SUBAPPLICATION logiBUS_AI_Calibrate_2P_IDA_Param_OPC (* logiBUS_AI_IDA (Analog-Eingang) mit 2-Punkt-Kalibrierung (AR_CALIBRATE_2P_REF, unabhaengig gespeicherte Rohwerte X_LOW/X_HIGH + Referenzwerte LOW_REF/HIGH_REF alle INI-persistiert) auf VT-Zahlenfelder (Rohwert + kalibrierter Wert, je eigene CNumberVariable) + Bargraph (kalibriert) + 2 VT-Tasten (CO/CS) + OPC-UA (Rohwert DWORD + kalibrierter Wert REAL, generisch, ein Kanal) *)
  (* Standard: 61499-2; Description: Copyright (c) 2026 Meisterschulen am Ostbahnhof This program and the accompanying materials are made available under the terms of the Eclipse Public License 2.0 which is available at https://www.eclipse.org/legal/epl-2.0/ SPDX-License-Identifier: EPL-2.0 *)
  (* Version 1.0, 2026-11-23, Franz Höpfinger, Meisterschulen am Ostbahnhof, Kopie von logiBUS_AI_Calibrate_2P_IDA_OPC (v1.13), InputRaw jetzt logiBUS_AI_Raw_VT_AR_Param_OPC: Hysterese/TimeDelta/TimeRateLimit des AI per Web + INI einstellbar (gleiche sSection). Zuerst fuer Ultraschall B01. PublishCal auf AR_TO_Q_Publish_Fast_OPC: CAL-Publish ungedrosselt, nur VT-Anzeige 500 ms. *)
  PACKAGE MyLib::sys;
  IMPORT isobus::UT::Q::const::IDs::ID_NULL;
  IMPORT logiBUS::io::AI::logiBUS_AI;
  IMPORT logiBUS::io::AI::logiBUS_AI_S;
  IMPORT logiBUS::utils::conversion::phys::NumericObjectPool_S;
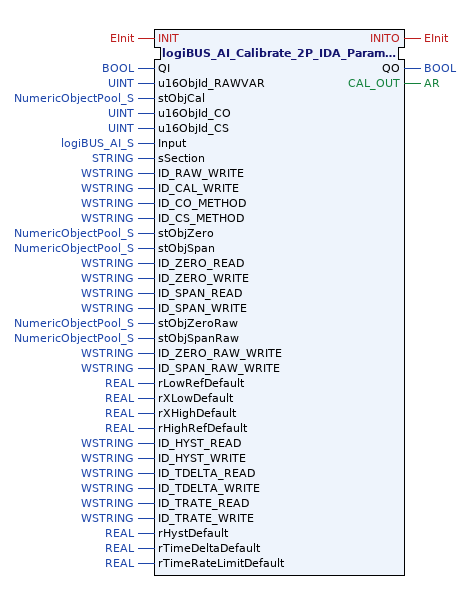
  EVENT_INPUT
    INIT : EInit; (* Initialization Request *)
  END_EVENT
  EVENT_OUTPUT
    INITO : EInit; (* Initialization Confirm *)
  END_EVENT
  VAR_INPUT
    QI : BOOL := TRUE; (* Quality Input - TRUE to enable service *)
    u16ObjId_RAWVAR : UINT := ID_NULL; (* Object ID CNumberVariable (Rohwert 0-4095, unkalibriert, reine Diagnose-Anzeige) *)
    stObjCal : logiBUS::utils::conversion::phys::NumericObjectPool_S := (u16ObjId := ID_NULL, r32Scale := 1.0, i32Offset := 0, u8Decimals := 1); (* Object ID + Scale/Offset/Decimals CNumberVariable (kalibrierter Wert, eigene, unabhaengige CNumberVariable) *)
    u16ObjId_CO : UINT := ID_NULL; (* Object ID Taste 'CO' (Kalibrier-Nullpunkt: Referenz 1 anlegen, dann druecken) *)
    u16ObjId_CS : UINT := ID_NULL; (* Object ID Taste 'CS' (Kalibrier-Spanne: Referenz 2 anlegen, dann druecken - erst nach CO moeglich) *)
    Input : logiBUS::io::AI::logiBUS_AI_S := logiBUS_AI::Invalid; (* Identify the Input AnalogInput_I1..I8 *)
    sSection : STRING; (* INI-Sektionsname fuer OFFSET/SCALE-Persistenz - pro Kanal eindeutig (z.B. 'AI_Calibrate_I1'), sonst kollidieren die Kanaele in settings.ini *)
    ID_RAW_WRITE : WSTRING; (* Rohwert-Ruckmelde-Adresse (DWORD 0-4095, ACTION=PUBLISH) *)
    ID_CAL_WRITE : WSTRING; (* Kalibrierter-Wert-Ruckmelde-Adresse (REAL, ACTION=PUBLISH) *)
    ID_CO_METHOD : WSTRING; (* Methodenadresse (ACTION=CREATE_METHOD) fuer den argumentlosen CO-Trigger - gleichberechtigt zur lokalen VT-Taste aufrufbar, sowohl vom OPC-UA-Dashboard als auch per CLIENT_0 von einer anderen Station (Cross-Station-Weiterleitung einer dortigen VT-Taste, siehe OPC_UA_VERNETZUNG.md Punkt 14 - kein Toggle/Subscribe-Umweg mehr) *)
    ID_CS_METHOD : WSTRING; (* Methodenadresse (ACTION=CREATE_METHOD) fuer den argumentlosen CS-Trigger - siehe ID_CO_METHOD *)
    stObjZero : logiBUS::utils::conversion::phys::NumericObjectPool_S := (u16ObjId := ID_NULL, r32Scale := 1.0, i32Offset := 0, u8Decimals := 1); (* Object ID + Scale/Offset/Decimals CNumberVariable (ZERO-Referenzwert, VT-Eingabefeld + OPC-UA) *)
    stObjSpan : logiBUS::utils::conversion::phys::NumericObjectPool_S := (u16ObjId := ID_NULL, r32Scale := 1.0, i32Offset := 0, u8Decimals := 1); (* Object ID + Scale/Offset/Decimals CNumberVariable (SPAN-Referenzwert, VT-Eingabefeld + OPC-UA) *)
    ID_ZERO_READ : WSTRING; (* Remote-Subscribe-Adresse ZERO-Referenzwert (REAL, ACTION=SUBSCRIBE) *)
    ID_ZERO_WRITE : WSTRING; (* Remote-Echo-Adresse ZERO-Referenzwert (REAL, ACTION=PUBLISH) *)
    ID_SPAN_READ : WSTRING; (* Remote-Subscribe-Adresse SPAN-Referenzwert (REAL, ACTION=SUBSCRIBE) *)
    ID_SPAN_WRITE : WSTRING; (* Remote-Echo-Adresse SPAN-Referenzwert (REAL, ACTION=PUBLISH) *)
    stObjZeroRaw : logiBUS::utils::conversion::phys::NumericObjectPool_S := (u16ObjId := ID_NULL, r32Scale := 1.0, i32Offset := 0, u8Decimals := 1); (* Object ID + Scale/Offset/Decimals CNumberVariable (Rohwert am ZERO-Kalibrierpunkt, reine Diagnose-Anzeige) *)
    stObjSpanRaw : logiBUS::utils::conversion::phys::NumericObjectPool_S := (u16ObjId := ID_NULL, r32Scale := 1.0, i32Offset := 0, u8Decimals := 1); (* Object ID + Scale/Offset/Decimals CNumberVariable (Rohwert am SPAN-Kalibrierpunkt, reine Diagnose-Anzeige) *)
    ID_ZERO_RAW_WRITE : WSTRING; (* Rohwert-am-ZERO-Kalibrierpunkt-Publish-Adresse (REAL, ACTION=PUBLISH) *)
    ID_SPAN_RAW_WRITE : WSTRING; (* Rohwert-am-SPAN-Kalibrierpunkt-Publish-Adresse (REAL, ACTION=PUBLISH) *)
    rLowRefDefault : REAL := REAL#0.0; (* Erstinbetriebnahme-Standardwert LOW_REF (INI_LOW_REF.DEFAULT_VALUE), bevor der Bediener selbst kalibriert - Fuellband/die meisten Sensoren: 0.0 *)
    rXLowDefault : REAL := REAL#0.0; (* Erstinbetriebnahme-Rohwert X_LOW (INI_X_LOW.DEFAULT_VALUE) *)
    rXHighDefault : REAL := REAL#0.0; (* Erstinbetriebnahme-Rohwert X_HIGH (INI_X_HIGH.DEFAULT_VALUE) *)
    rHighRefDefault : REAL := REAL#100.0; (* Erstinbetriebnahme-Standardwert HIGH_REF (INI_HIGH_REF.DEFAULT_VALUE), bevor der Bediener selbst kalibriert - z.B. 250.0 fuer Druck (0-250bar), 100.0 fuer Fuellband-Winkel (Prozent) *)
    ID_HYST_READ : WSTRING; (* Web-Override AI-Hysterese (Digits) *)
    ID_HYST_WRITE : WSTRING; (* Rueckmeldung AI-Hysterese *)
    ID_TDELTA_READ : WSTRING; (* Web-Override AI-TimeDelta (ms) *)
    ID_TDELTA_WRITE : WSTRING; (* Rueckmeldung AI-TimeDelta *)
    ID_TRATE_READ : WSTRING; (* Web-Override AI-TimeRateLimit (ms) *)
    ID_TRATE_WRITE : WSTRING; (* Rueckmeldung AI-TimeRateLimit *)
    rHystDefault : REAL := 3.0; (* Default AI-Hysterese (Digits) *)
    rTimeDeltaDefault : REAL := 100.0; (* Default AI-TimeDelta (ms) *)
    rTimeRateLimitDefault : REAL := 20.0; (* Default AI-TimeRateLimit (ms) *)
  END_VAR
  VAR_OUTPUT
    QO : BOOL; (* Quality Output - TRUE if service executed successfully *)
  END_VAR
  PLUGS
    CAL_OUT : adapter::types::unidirectional::AR; (* Kalibrierter Wert, lokal (= CALIBRATE.Y) - fuer Weiterverarbeitung auf derselben Station ohne OPC-UA-Roundtrip *)
  END_PLUGS
  FBS
    CALIBRATE : adapter::Engineering::measurements::AR_CALIBRATE_2P_REF(xClipping := FALSE);
    INI_X_LOW : eclipse4diac::storage::INI_AR2(SETM := TRUE, KEY := 'X_LOW');
    INI_X_HIGH : eclipse4diac::storage::INI_AR2(SETM := TRUE, KEY := 'X_HIGH');
    INI_LOW_REF : eclipse4diac::storage::INI_AR2(SETM := TRUE, KEY := 'LOW_REF');
    INI_HIGH_REF : eclipse4diac::storage::INI_AR2(SETM := TRUE, KEY := 'HIGH_REF');
    TapZeroRaw : adapter::events::bidirectional::AR2_SPLIT_FWD_REV;
    TapSpanRaw : adapter::events::bidirectional::AR2_SPLIT_FWD_REV;
    AR_SPLIT_2_Cal : adapter::events::unidirectional::AR_SPLIT_2;
    AND_QO : iec61131::booleanOperators::AND_BOOL_13;
  END_FBS
  SUBAPPS
    InputRaw : MyLib::sys::logiBUS_AI_Raw_VT_AR_Param_OPC;
    Y_OFFSET_LIT : MyLib::sys::NumericValue_TO_AR2_OPC;
    Y_SCALE_LIT : MyLib::sys::NumericValue_TO_AR2_OPC;
    TriggerCO : MyLib::sys::Button_Method_IE;
    TriggerCS : MyLib::sys::Button_Method_IE;
    PublishCal : MyLib::sys::AR_TO_Q_Publish_Fast_OPC;
    PublishZeroRaw : MyLib::sys::AR_TO_Q_Publish_OPC;
    PublishSpanRaw : MyLib::sys::AR_TO_Q_Publish_OPC;
  END_SUBAPPS
  EVENT_CONNECTIONS
    TriggerCO.IND TO CALIBRATE.C_LOW;
    TriggerCS.IND TO CALIBRATE.C_HIGH;
    INIT TO CALIBRATE.INIT;
    CALIBRATE.INITO TO INI_X_LOW.INIT;
    INI_X_LOW.INITO TO INI_X_HIGH.INIT;
    INI_X_HIGH.INITO TO INI_LOW_REF.INIT;
    INI_LOW_REF.INITO TO INI_HIGH_REF.INIT;
    INI_HIGH_REF.INITO TO InputRaw.INIT;
    InputRaw.INITO TO Y_OFFSET_LIT.INIT;
    Y_OFFSET_LIT.INITO TO Y_SCALE_LIT.INIT;
    Y_SCALE_LIT.INITO TO TriggerCO.INIT;
    TriggerCO.INITO TO TriggerCS.INIT;
    TriggerCS.INITO TO PublishCal.INIT;
    PublishCal.INITO TO PublishZeroRaw.INIT;
    PublishZeroRaw.INITO TO PublishSpanRaw.INIT;
    PublishSpanRaw.INITO TO INITO;
    PublishSpanRaw.INITO TO AND_QO.REQ;
  END_CONNECTIONS
  DATA_CONNECTIONS
    rXLowDefault TO INI_X_LOW.DEFAULT_VALUE;
    rXHighDefault TO INI_X_HIGH.DEFAULT_VALUE;
    Input TO InputRaw.Input;
    u16ObjId_RAWVAR TO InputRaw.u16ObjId_RAWVAR;
    stObjCal TO PublishCal.stObj;
    u16ObjId_CO TO TriggerCO.u16ObjId;
    u16ObjId_CS TO TriggerCS.u16ObjId;
    sSection TO INI_X_LOW.SECTION;
    sSection TO INI_X_HIGH.SECTION;
    sSection TO INI_LOW_REF.SECTION;
    sSection TO INI_HIGH_REF.SECTION;
    rLowRefDefault TO INI_LOW_REF.DEFAULT_VALUE;
    rHighRefDefault TO INI_HIGH_REF.DEFAULT_VALUE;
    ID_RAW_WRITE TO InputRaw.ID_RAW_WRITE;
    ID_CAL_WRITE TO PublishCal.ID_WRITE;
    ID_CO_METHOD TO TriggerCO.ID_METHOD;
    ID_CS_METHOD TO TriggerCS.ID_METHOD;
    stObjZero TO Y_OFFSET_LIT.stObj;
    ID_ZERO_READ TO Y_OFFSET_LIT.ID_READ;
    ID_ZERO_WRITE TO Y_OFFSET_LIT.ID_WRITE;
    stObjSpan TO Y_SCALE_LIT.stObj;
    ID_SPAN_READ TO Y_SCALE_LIT.ID_READ;
    ID_SPAN_WRITE TO Y_SCALE_LIT.ID_WRITE;
    stObjZeroRaw TO PublishZeroRaw.stObj;
    ID_ZERO_RAW_WRITE TO PublishZeroRaw.ID_WRITE;
    stObjSpanRaw TO PublishSpanRaw.stObj;
    ID_SPAN_RAW_WRITE TO PublishSpanRaw.ID_WRITE;
    QI TO CALIBRATE.QI;
    QI TO INI_X_LOW.QI;
    QI TO INI_X_HIGH.QI;
    QI TO INI_LOW_REF.QI;
    QI TO INI_HIGH_REF.QI;
    QI TO InputRaw.QI;
    QI TO Y_OFFSET_LIT.QI;
    QI TO Y_SCALE_LIT.QI;
    QI TO TriggerCO.QI;
    QI TO TriggerCS.QI;
    QI TO PublishCal.QI;
    QI TO PublishZeroRaw.QI;
    QI TO PublishSpanRaw.QI;
    CALIBRATE.QO TO AND_QO.IN1;
    INI_X_LOW.QO TO AND_QO.IN2;
    INI_X_HIGH.QO TO AND_QO.IN3;
    INI_LOW_REF.QO TO AND_QO.IN4;
    INI_HIGH_REF.QO TO AND_QO.IN5;
    InputRaw.QO TO AND_QO.IN6;
    Y_OFFSET_LIT.QO TO AND_QO.IN7;
    Y_SCALE_LIT.QO TO AND_QO.IN8;
    TriggerCO.QO TO AND_QO.IN9;
    TriggerCS.QO TO AND_QO.IN10;
    PublishCal.QO TO AND_QO.IN11;
    PublishZeroRaw.QO TO AND_QO.IN12;
    PublishSpanRaw.QO TO AND_QO.IN13;
    AND_QO.OUT TO QO;
    sSection TO InputRaw.sSection;
    ID_HYST_READ TO InputRaw.ID_HYST_READ;
    ID_HYST_WRITE TO InputRaw.ID_HYST_WRITE;
    ID_TDELTA_READ TO InputRaw.ID_TDELTA_READ;
    ID_TDELTA_WRITE TO InputRaw.ID_TDELTA_WRITE;
    ID_TRATE_READ TO InputRaw.ID_TRATE_READ;
    ID_TRATE_WRITE TO InputRaw.ID_TRATE_WRITE;
    rHystDefault TO InputRaw.rHystDefault;
    rTimeDeltaDefault TO InputRaw.rTimeDeltaDefault;
    rTimeRateLimitDefault TO InputRaw.rTimeRateLimitDefault;
  END_CONNECTIONS
  ADAPTER_CONNECTIONS
    InputRaw.AR_OUT TO CALIBRATE.X;
    CALIBRATE.X_LOW TO TapZeroRaw.IN;
    TapZeroRaw.OUT TO INI_X_LOW.VAL;
    TapZeroRaw.REV_OUT TO PublishZeroRaw.AR_IN;
    CALIBRATE.X_HIGH TO TapSpanRaw.IN;
    TapSpanRaw.OUT TO INI_X_HIGH.VAL;
    TapSpanRaw.REV_OUT TO PublishSpanRaw.AR_IN;
    CALIBRATE.LOW_REF TO INI_LOW_REF.VAL;
    CALIBRATE.HIGH_REF TO INI_HIGH_REF.VAL;
    Y_OFFSET_LIT.VALUEO TO CALIBRATE.Y_LOW;
    Y_SCALE_LIT.VALUEO TO CALIBRATE.Y_HIGH;
    CALIBRATE.Y TO AR_SPLIT_2_Cal.IN;
    AR_SPLIT_2_Cal.OUT2 TO PublishCal.AR_IN;
    AR_SPLIT_2_Cal.OUT1 TO CAL_OUT;
  END_CONNECTIONS
END_SUBAPPLICATION
